        - object Box at (437051, 103.35, 13.17) mm, rotated rx -0.53 ry 0.26 rz 8.05 deg, size 10 x 20 x 5 mm, geometry from box.sld
        - object Box at (436264, 103.35, 13.17) mm, rotated rx -0.42 ry 0.42 rz 26.92 deg, size 10 x 20 x 5 mm, geometry from box.sld
        - object Box at (435475, 103.35, 13.17) mm, rotated rx -0.46 ry 0.37 rz 20.31 deg, size 10 x 20 x 5 mm, geometry from box.sld
        - object Box at (434685, 103.35, 13.17) mm, rotated rx -0.45 ry 0.39 rz 22.66 deg, size 10 x 20 x 5 mm, geometry from box.sld
        - object Box at (433900, 103.35, 13.17) mm, rotated rx -0.59 ry 0.03 rz -15.41 deg, size 10 x 20 x 5 mm, geometry from box.sld
        - object Box at (433098, 103.35, 13.17) mm, rotated rx -0.53 ry 0.28 rz 9.45 deg, size 10 x 20 x 5 mm, geometry from box.sld
    - frame Reference Box Frame at (60, 290, 366.5) mm
      - object ref_obj at (0, 0, 0) mm, size 252 x 305.4 x 216.7 mm, geometry from Box-12x10in-Closed.sld
      - object ref_lid at (-60, -186.65, 13.17) mm, rotated rx -0.56 ry 0.19 rz 0 deg, size 10 x 20 x 5 mm, geometry from box.sld
    - object SICK WL4S Laser Sensor at (1954, -20, 370) mm, rotated rx 180 ry 0 rz 90 deg, size 683.3 x 45.2 x 12.5 mm, geometry from SICK-WL4S-Laser-Sensor.sld
    - object start_prox at (0, -20, 370) mm, rotated rx 180 ry 0 rz 90 deg, size 683.3 x 45.2 x 12.5 mm, geometry from SICK-WL4S-Laser-Sensor.sld
